(* PLC project TBEN_L5_PLC11.project, CODESYS CODESYS V3.5 SP21 Patch 1 *)
(* stored: creationDateTime 2026-11-07T15:34:51.1476266, modificationDateTime 2026-11-07T15:09:07.4034196 *)

{attribute 'qualified_only'}
// Bước trình tự gọi ISDU trong FB_IolDevBase
TYPE E_IolDevSeq :
(
    IDLE    := 0,   // chọn việc tiếp theo
    RUN     := 1,   // FB_IolCall đang chạy
    RELEASE := 2    // hạ Execute, chờ FB_IolCall về IDLE
) INT;
END_TYPE
